(* IEC 61131-3 sources: plc-workbench/outputs/tia_32x4_20261108_results/tasks/02_CUSTOM_02/self_B/details/submissions/2/evaluation/formal, 1 file *)

(* ---- normalized.st ---- *)
FUNCTION_BLOCK FB_HmiAccess

VAR_INPUT
    SessionValid : BOOL;
    Role : USINT;
    Page : USINT;
    WriteReq : BOOL;
    WriteValue : LREAL;
END_VAR

VAR_OUTPUT
    ViewAllowed : BOOL;
    WriteAllowed : BOOL;
    Accepted : BOOL;
    Denied : BOOL;
    ParamValue : LREAL;
END_VAR

VAR_IN_OUT
END_VAR

VAR
    m_ParamValue : LREAL := 0.0;
END_VAR

VAR
    t_IsAuthorizedUser : BOOL;
    t_CanViewPage : BOOL;
    t_ValueInRange : BOOL;
END_VAR
VAR_INPUT
WBTEMP_0 : BOOL;
WBTEMP_1 : BOOL;
WBTEMP_2 : BOOL;
END_VAR

t_IsAuthorizedUser := WBTEMP_0;
t_CanViewPage := WBTEMP_1;
t_ValueInRange := WBTEMP_2;
    // Initialize outputs for current scan
    Accepted := FALSE;
    Denied := FALSE;

    // Determine if the role is valid (1=user, 2=operator, 3=admin)
    t_IsAuthorizedUser := (Role = 1) OR (Role = 2) OR (Role = 3);

    // Calculate ViewAllowed based on requirements:
    // Admin (3): Pages 1..4
    // Operator (2): Pages 1, 2, 4
    // User (1): Pages 1, 2
    IF SessionValid AND t_IsAuthorizedUser THEN
        CASE Role OF
            1: // User
                t_CanViewPage := (Page = 1) OR (Page = 2);
            2: // Operator
                t_CanViewPage := (Page = 1) OR (Page = 2) OR (Page = 4);
            3: // Administrator
                t_CanViewPage := (Page >= 1) AND (Page <= 4);
            ELSE
                t_CanViewPage := FALSE;
        END_CASE;
    ELSE
        t_CanViewPage := FALSE;
    END_IF;

    ViewAllowed := t_CanViewPage;

    // Calculate WriteAllowed:
    // TRUE only for Page 4 with valid session and Role 2 or 3
    WriteAllowed := SessionValid AND ((Role = 2) OR (Role = 3)) AND (Page = 4);

    // Handle Parameter Write Request
    IF WriteReq THEN
        IF WriteAllowed THEN
            // Check if value is in range [0, 100]
            t_ValueInRange := (WriteValue >= 0.0) AND (WriteValue <= 100.0);

            IF t_ValueInRange THEN
                // Accept the write
                m_ParamValue := WriteValue;
                Accepted := TRUE;
                Denied := FALSE;
            ELSE
                // Reject due to out-of-range value
                Accepted := FALSE;
                Denied := TRUE;
            END_IF;
        ELSE
            // Reject due to insufficient permission
            Accepted := FALSE;
            Denied := TRUE;
        END_IF;
    ELSE
        // No request made
        Accepted := FALSE;
        Denied := FALSE;
    END_IF;

    // Update output parameter with retained state
    ParamValue := m_ParamValue;

END_FUNCTION_BLOCK
